(* IEC 61131-3 sources: trust-platform/examples/blockly, 2 files *)

(* ---- snake-simple-v2.st ---- *)
(*
  Auto-generated from blockly source: snake-simple-v2.blockly.json
  Source of truth is the visual file unless migrated fully to ST.
*)
(*
  Blockly conversion warnings (1):
  - Unknown block type: controls_whileUntil
*)

FUNCTION_BLOCK FB_snake_simple_v2_BLOCKLY

VAR
  position : BOOL;
  direction : BOOL;
  temp : INT;
END_VAR

(* Generated from Blockly *)

temp := 0;
temp := 1;
(* Unknown block: controls_whileUntil *)

END_FUNCTION_BLOCK

(* ---- snake-simple-v2.visual.runtime.st ---- *)
(*
  Auto-generated runtime entry for snake-simple-v2.blockly.json.
  This wrapper is used to run visual editors through the Structured Text debugger path.
*)

PROGRAM PRG_snake_simple_v2_VISUAL
fb_snake_simple_v2();
END_PROGRAM

CONFIGURATION CFG_snake_simple_v2_VISUAL
VAR_GLOBAL
  fb_snake_simple_v2 : FB_snake_simple_v2_BLOCKLY;
END_VAR
  RESOURCE RES_snake_simple_v2_VISUAL ON PLC
    TASK TASK_snake_simple_v2_VISUAL(INTERVAL := T#20ms, PRIORITY := 1);
    PROGRAM PLC_PRG_snake_simple_v2 WITH TASK_snake_simple_v2_VISUAL : PRG_snake_simple_v2_VISUAL;
  END_RESOURCE
END_CONFIGURATION
